Fanuc KAREL source: kt00441.KL

-- PROVISIONAL review KL for V940-1; original PC SHA256 ff04b8d79f561274b954aa898d406792c01a4d259d6860ab46bd4cc085f33c5c
-- Incomplete behavior may be omitted. Consult companion uncertainty JSON. Do not deploy.
PROGRAM KT00441
%NOLOCKGROUP
VAR
  R1 : REAL
  I2 : INTEGER
  OUT : BOOLEAN
BEGIN
  -- V9_ZERO_TABLE_METADATA_HINT layout=0001; no indexed target words; source/name/runtime held
  -- UNRESOLVED_PC offsets 5-16; opcodes 2E,23
  -- UNRESOLVED_PC offsets 21-32; opcodes 2E,23
  -- UNRESOLVED_PC offsets 37-57; opcodes 21,21,64,72,23
  -- UNRESOLVED_PC offsets 62-66; opcodes 7F
END KT00441
